Fanuc KAREL source: kt00552.KL

-- PROVISIONAL review KL for V940-1; original PC SHA256 c1cfdeb5679ade50983746514c7b767230ee8f82355dd96b5df85b45c4c3d345
-- Incomplete behavior may be omitted. Consult companion uncertainty JSON. Do not deploy.
PROGRAM KT00552
%NOLOCKGROUP
-- UNRESOLVED_DECL P1 type=000199
-- UNRESOLVED_DECL P2 type=000199
-- UNRESOLVED_DECL OUT type=000199
BEGIN
  -- V9_ZERO_TABLE_METADATA_HINT layout=0001; no indexed target words; source/name/runtime held
  -- UNRESOLVED_PC offsets 5-44; opcodes 49,7E,49,7E,60,7E,4A
  -- UNRESOLVED_PC offsets 49-53; opcodes 7F
END KT00552
